// TIA Portal V21 export
// export: Created 2026-11-11T00:47:41.9876793Z, ExportSetting WithDefaults, DisplayName Totally Integrated Automation Portal, DisplayVersion V21 Update 3, DisplayName STEP 7 Professional, DisplayVersion V21 Update 3, DisplayName STEP 7 Safety, DisplayVersion V21, DisplayName Tech WebApplication, DisplayVersion V21, DisplayName WinCC Basic/Comfort/Advanced, DisplayVersion V21 Update 3, DisplayName WinCC Unified, DisplayVersion V21 Update 3
FUNCTION_BLOCK "FB_Fbd_ex158"   // FB166, FBD
{ S7_Optimized_Access := 'TRUE' }
VERSION : 0.1
// stored: AutoNumber true, IsIECCheckEnabled false, IsRetainMemResEnabled false, MemoryReserve 100, SetENOAutomatically false, UDAEnableTagReadback false
   VAR_INPUT
      v_laddr : HW_IO;
   END_VAR
   VAR_OUTPUT
      v_ret_val : Int;
      v_area : Int;
      v_master : Int;
      v_station : Int;
      v_slot : Int;
      v_subslot : Int;
      v_offset : Int;
   END_VAR
BEGIN

REGION Network 1: LOG_GEO - Determine slot from hardware identifier
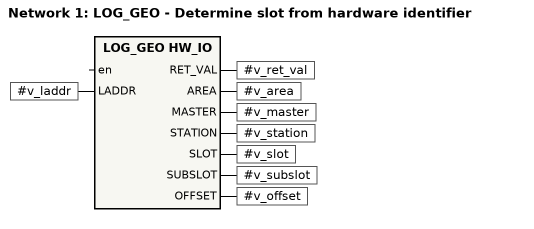
   #v_ret_val := LOG_GEO(LADDR := #v_laddr,
                         AREA => #v_area,
                         MASTER => #v_master,
                         STATION => #v_station,
                         SLOT => #v_slot,
                         SUBSLOT => #v_subslot,
                         OFFSET => #v_offset);
END_REGION
END_FUNCTION_BLOCK
